Fanuc KAREL source: kt00038.KL

-- PROVISIONAL review KL for V1013-1; original PC SHA256 630a878c6e4d22fecdef786c9591a44dbd75317392d2e83b49d8884bf5c68f66
-- Incomplete behavior may be omitted. Consult companion uncertainty JSON. Do not deploy.
PROGRAM KT00038
%NOLOCKGROUP
VAR
  I1 : INTEGER
  OUT : REAL
-- UNRESOLVED_DECL Y2 type=002018
BEGIN
  -- UNRESOLVED_PC offsets 5-16; opcodes 2E,23
  -- UNRESOLVED_PC offsets 21-35; opcodes 2E,22,9D,33,B2
  -- UNRESOLVED_PC offsets 40-63; opcodes 21,22,9D,33,B1,53,64,23
  -- UNRESOLVED_PC offsets 68-72; opcodes 7F
END KT00038
